Fanuc KAREL source: KC00025.KL

PROGRAM KC00025
%NOLOCKGROUP
%ENVIRONMENT UIF
VAR
  I: INTEGER
  J: INTEGER
  K: INTEGER
  R: REAL
  B: BOOLEAN
  S: STRING[80]
  T: STRING[80]
  P: PATH
  Q: PATH
  AI: ARRAY[8] OF INTEGER
  AB: ARRAY[244] OF BYTE
BEGIN
  S = 'DICT'
  DISCTRL_PLMN(S,I,J,K,I,J)
END KC00025
